(* PLC project Vn_return_uncond, Beckhoff Automation GmbH TwinCAT PLC Control 3.5.13.21 *)
(* stored: creationDateTime 1970-01-01T00:00:00 *)

PROGRAM Vn_return_uncond

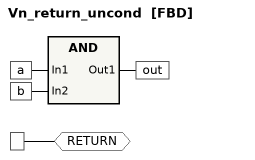
(* FBD diagram, written out as Structured Text *)
out := a AND b;
IF  THEN RETURN; END_IF;
END_PROGRAM
